// TIA Portal V20 export
// export: Created 2026-10-19T18:02:43.4272931Z, ExportSetting WithDefaults, DisplayName Totally Integrated Automation Portal, DisplayVersion V20 Update 6, DisplayName TIA Portal Openness, DisplayVersion V20 Update 6, DisplayName TIA Portal Version Control Interface, DisplayVersion V20 Update 6, DisplayName SINAMICS Startdrive Advanced, DisplayVersion V20 SP1, DisplayName SINAMICS Startdrive G130, G150, S120, S150, SINAMICS MV, G220, S200, S210, DisplayVersion V20 SP1, DisplayName SINAMICS Startdrive G110M, G120, G120C, G120D, G120P, G115D, DisplayVersion V20 SP1, DisplayName STEP 7 Professional, DisplayVersion V20 Update 6, DisplayName STEP 7 Safety, DisplayVersion V20 Update 2, DisplayName WinCC Basic/Comfort/Advanced, DisplayVersion V20 Update 6, DisplayName WinCC Unified, DisplayVersion V20 Update 6
DATA_BLOCK "OPC_UA_Control_FB_DB"   // DB17
VERSION : 0.1
// stored: AutoNumber true, DBAccessibleFromOPCUA true, DBAccessibleFromWebserver true, InstanceOfName OPC_UA_Control_FB, InstanceOfType FB
"OPC_UA_Control_FB"
   // VAR_INPUT
   //    OPC_Enable : Bool;
   //    Mode_Change : UInt;
   // END_VAR
   // VAR_OUTPUT
   //    Mode_Current : UInt;
   // END_VAR
   // VAR
   //    Source_Location_VTD { ExternalAccessible := 'False'; ExternalVisible := 'False'; ExternalWritable := 'False'} : "ID_Decoded";
   //    Destination_Location_VTD { ExternalAccessible := 'False'; ExternalVisible := 'False'; ExternalWritable := 'False'} : "ID_Decoded";
   //    Source_Location_Carousel { ExternalAccessible := 'False'; ExternalVisible := 'False'; ExternalWritable := 'False'} : "ID_Decoded";
   //    Destination_Location_Carousel { ExternalAccessible := 'False'; ExternalVisible := 'False'; ExternalWritable := 'False'} : "ID_Decoded";
   //    State_VTD : UInt;
   //    State_Carrousel_Weigh : UInt;
   //    State_Carrousel_Main : UInt;
   //    State_Carrousel_PICKTP1 : UInt;
   //    State_Carrousel_P4TPICK : UInt;
   //    State_Carrousel_CTC : UInt;
   //    State_Carrousel_ITP1 : UInt;
   //    State_Carrousel_P1TP2 : UInt;
   //    State_Carrousel_P3TP4 : UInt;
   //    State_Carrousel_P4TO : UInt;
   //    State_Carrousel : UInt;
   // END_VAR
BEGIN
END_DATA_BLOCK
